PROGRAM ladder
VAR
	xoutput: BOOL;
	xtest: BOOL;
	xtest2: BOOL;
END_VAR
VAR // added by the converter: edge detectors and wires of the graphical bodies
    _w1 : BOOL;
END_VAR

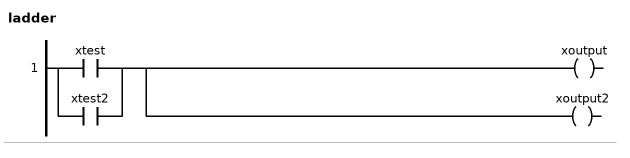
// NETWORK 1
_w1 := xtest OR xtest2;
xoutput := _w1;
xoutput2 := _w1;

END_PROGRAM

(* stored: Version 1.1.0.1, ProductVersion 3.1.4024.16
   POU ladder: Id {04d867c5-831f-4a2c-a8ba-57738ccf38e1}, SpecialFunc None *)
